    rq_activate_all_grippers(True)
    # end: URCap Program Node
  end
  $ 60 "zero_ftsensor()"
  zero_ftsensor()
  $ 61 "EXTT"
  $ 62 "Set GRP_3F_Enable=Off"
  set_standard_digital_out(4, False)
  $ 63 "Set BarcodeTrigger=Off"
  set_standard_digital_out(6, False)
  $ 64 "Set GRP_3F_Decap=Off"
  set_standard_digital_out(3, False)
  $ 65 "Set GRP_3F_Cap=Off"
  set_standard_digital_out(2, False)
  $ 66 "Set GRP_3F_Open=Off"
  set_standard_digital_out(5, False)
  $ 67 "PSE_T≔get_tool_free_pose(dir=[0,0,0.150], move_in_base_frame=True)"
  global PSE_T=get_tool_free_pose(dir=[0,0,0.150], move_in_base_frame=True)
  $ 68 "If is_reachable(Base_const, [PSE_T])"
  if (is_reachable(p[0.0,0.0,0.0,0.0,0.0,0.0], [PSE_T])):
    $ 69 "MoveL"
    $ 70 "PSE_T" "breakAfter"
    movel(PSE_T, a=1.2, v=0.15)
  end
  $ 71 "powder dispensing variable init"
  $ 72 "Start_thread≔ False "
  global Start_thread=  False
  $ 73 "vib_thread≔ False "
  global vib_thread=  False
  $ 74 "kp≔0.0015"
  global kp=0.0015
  $ 75 "ki≔0.0001"
  global ki=0.0001
  $ 76 "kd≔0.01"
  global kd=0.01
  $ 77 "dt≔0.03"
  global dt=0.03
  $ 78 "Integral_error≔0"
  global Integral_error=0
  $ 79 "current_error≔0"
  global current_error=0
  $ 80 "previous_error≔0"
  global previous_error=0
  $ 81 "tilt_increment≔0"
  global tilt_increment=0
  $ 82 "tilt_angle≔0"
  global tilt_angle=0
  $ 83 "diff≔0"
  global diff=0
  $ 84 "current_pose≔get_actual_tcp_pose()"
  global current_pose= get_actual_tcp_pose ()
  $ 85 "Relative_trans≔p[0, 0, -0.035, 0, 0, 0]"
  global Relative_trans=p[0, 0, -0.035, 0, 0, 0]
  $ 86 "ContA_plc_offst≔p[-0.00205, 0.02547, 0.03730, -0.03, -2.183, 6.165]"
  global ContA_plc_offst=p[-0.00205, 0.02547, 0.03730, -0.03, -2.183, 6.165]
  $ 87 "PowA_50_offset≔p[0.21808, -0.19943, 0.06584, 0, 0, 0]"
  global PowA_50_offset=p[0.21808, -0.19943, 0.06584, 0, 0, 0]
  $ 89 "tilt_init_reference()"
  tilt_init_reference()
  $ 90 "switch_spat_M≔ True "
  global switch_spat_M=  True
  $ 91 "switch_spat_S≔ True "
  global switch_spat_S=  True
  $ 92 "switch_spat_F_M≔ True "
  global switch_spat_F_M=  True
  $ 93 "switch_spat_F_S≔ True "
  global switch_spat_F_S=  True
  $ 94 "last_scale≔0"
  global last_scale=0
  $ 95 "W_EMPTY≔51.3"
  global W_EMPTY=51.3
  $ 768 "Thread_1"
  thread Thread_1():
    while (True):
      $ 769 "If Start_thread≟ True "
      if (Start_thread ==   True  ):
        $ 770 "weight_value≔get_weight()"
        global weight_value=get_weight()
        $ 771 "Wait: 0.1"
        sleep(0.1)
        $ 772 "sync()"
        sync()
      end
      $ 773 "sync()"
      sync()
    end
  end
  threadId_Thread_1 = run Thread_1()
  $ 774 "Thread_2"
  thread Thread_2():
    while (True):
      $ 775 "Loop vib_thread≟ True "
      thread Thread_while_775():
        while (True):
          $ 776 "diff≔target_weight-weight_value"
          global diff=target_weight-weight_value
          $ 777 "If diff>0.02 and spatula≠'spatula_flat_S'"
          global thread_flag_777=0
          thread Thread_if_777():
            $ 779 "Set AO[0]=4.0"
            set_standard_analog_out(0, 0.4)
            thread_flag_777 = 1
          end
          if (diff>0.02  and  spatula != "spatula_flat_S"):
            global thread_handler_777=run Thread_if_777()
            while (thread_flag_777 == 0):
              if not(diff>0.02  and  spatula != "spatula_flat_S"):
                kill thread_handler_777
                thread_flag_777 = 2
              else:
                sync()
              end
            end
          else:
            thread_flag_777 = 2
          end
          if (thread_flag_777 == 2):
            $ 780 "ElseIf diff>0.02 and spatula≟'spatula_flat_S'"
            if (diff>0.02 and spatula == "spatula_flat_S"):
              $ 781 "vibration_3()"
              vibration_3()
            else:
              $ 782 "ElseIf diff≤0.03"
              global thread_flag_782=0
              thread Thread_if_782():
                $ 783 "vibration_2()"
                vibration_2()
                thread_flag_782 = 1
              end
              if (diff <= 0.03):
                global thread_handler_782=run Thread_if_782()
                while (thread_flag_782 == 0):
                  if not(diff <= 0.03):
                    kill thread_handler_782
                    thread_flag_782 = 2
                  else:
                    sync()
                  end
                end
              else:
                thread_flag_782 = 2
              end
              if (thread_flag_782 == 2):
                $ 788 "Else" "noBreak"
                $ 789 "Set AO[0]=0.0"
                set_standard_analog_out(0, 0.0)
              end
            end
          end
        end
      end
      if (vib_thread ==   True  ):
        global thread_handler_775=run Thread_while_775()
        while (vib_thread ==   True  ):
          sync()
        end
        kill thread_handler_775
      end
      $ 790 "sync()"
      sync()
    end
  end
  threadId_Thread_2 = run Thread_2()
  while (True):
    $ 96 "Robot Program"
    $ 97 "MAIN"
    $ 98 "command_manager(external_control='uGO', cond_suspend=(ITM_Manipulated and AMR_AtTarget and AMR_Charging and AMR_Battery<40), cond_unsuspend=(AMR_Battery≟60))"
    command_manager(external_control="uGO", cond_suspend=(ITM_Manipulated  and  AMR_AtTarget  and  AMR_Charging  and  AMR_Battery<40), cond_unsuspend=(AMR_Battery == 60))
    $ 99 "log_state(STATE_Info)"
    log_state(STATE_Info)
    $ 100 "Switch STATE"
    switch_1 = STATE
    $ 101 "Case 1"
    if (1 == switch_1):
      $ 102 "Stopping"
      $ 103 "STATE_Info≔'Stopping'"
      global STATE_Info="Stopping"
      $ 104 "end_freedrive_mode()"
      end_freedrive_mode()
      $ 105 "Set"
      set_tcp(p[0.0,0.0,0.161,3.1415,0.0,0.0])
      $ 106 "PSE_T≔get_tool_free_pose(dir=[0,0,0.150], move_in_base_frame=True)"
      global PSE_T=get_tool_free_pose(dir=[0,0,0.150], move_in_base_frame=True)
      $ 107 "If is_reachable(Base_const, [PSE_T])"
      if (is_reachable(p[0.0,0.0,0.0,0.0,0.0,0.0], [PSE_T])):
        $ 108 "MoveL"
        $ 109 "PSE_T" "breakAfter"
        movel(PSE_T, a=1.2, v=0.15)
      end
      $ 110 "do_transition(keep_rxry=OBJ_Picked, r=0)"
      do_transition(keep_rxry=OBJ_Picked, r=0)
      $ 119 "Call Sub_AMR_MiR_V3"
      Sub_AMR_MiR_V3()
      $ 120 "If stopping() and AMR_Done"
      if (stopping()  and  AMR_Done):
        $ 121 "STATE≔2"
        global STATE=2
        $ 122 "ugo_update_outputs()"
        ugo_update_outputs()
      end
    elif (2 == switch_1):
      $ 123 "Case 2"
      $ 124 "Stopped"
      $ 125 "STATE_Info≔'Stopped'"
      global STATE_Info="Stopped"
      $ 126 "Call Sub_AMR_MiR_V3"
      Sub_AMR_MiR_V3()
      $ 127 "If CMD_Reset  or PB_Start"
      if (CMD_Reset   or  get_standard_digital_in(0)):
        $ 128 "STATE≔3"
        global STATE=3
        $ 129 "ugo_update_outputs()"
        ugo_update_outputs()
      end
    elif (3 == switch_1):
      $ 130 "Case 3"
      $ 131 " Resetting"
      $ 132 "STATE_Info≔'Resetting'"
      global STATE_Info="Resetting"
      $ 133 "uML"
      $ 134 "reset_error()"
      reset_error()
      $ 135 "reset_warning()"
      reset_warning()
      $ 136 "PROCESS_Step≔0"
      global PROCESS_Step=0
      $ 137 "PROCESS_Info≔''"
      global PROCESS_Info=""
      $ 138 "ARM_Referenced≔ False "
      global ARM_Referenced=  False
      $ 139 "WRK_Done≔ False "
      global WRK_Done=  False
      $ 140 "ITM_Prepared≔ False "
      global ITM_Prepared=  False
      $ 141 "ITM_Manipulated≔ False "
      global ITM_Manipulated=  False
      $ 142 "STP≔0"
      global STP=0
      $ 143 "Action≔0"
      global Action=0
      $ 144 "Action_Info≔''"
      global Action_Info=""
      $ 145 "ITM_ID≔0"
      global ITM_ID=0
      $ 146 "JIG≔0"
      global JIG=0
      $ 147 "JIG_Slot≔0"
      global JIG_Slot=0
      $ 148 "Task_info≔''"
      global Task_info=""
      $ 149 "Set"
      set_tcp(p[0.0,0.0,0.161,3.1415,0.0,0.0])
      $ 150 "App"
      $ 151 "'ADD APPLICATION SPECIFIC COMMANDS'"
      # 'ADD APPLICATION SPECIFIC COMMANDS'
      $ 152 "OBJ_Type≔0"
      global OBJ_Type=0
      $ 153 "OBJ_Nbr≔0"
      global OBJ_Nbr=0
      $ 154 "If CNT_Rack_Output≥50"
      if (CNT_Rack_Output >= 50):
        $ 155 "CNT_Rack_Output≔0"
        global CNT_Rack_Output=0
      end
      $ 156 "TASK≔struct(ID=0, NAVI=struct(target=0, footprint=0, protectiveOff=0, dock=0), WORK=struct(ITM_ID_Src=0, JIG_ID_Src=0, OBJ_Nbr_Src=0, ACT_Src=0, ITM_ID_Tgt=0, JIG_ID_Tgt=0, OBJ_Nbr_Tgt=0, ACT_Tgt=0, OBJ_Type=0))"
      global TASK=struct(ID=0, NAVI=struct(target=0, footprint=0, protectiveOff=0, dock=0), WORK=struct(ITM_ID_Src=0, JIG_ID_Src=0, OBJ_Nbr_Src=0, ACT_Src=0, ITM_ID_Tgt=0, JIG_ID_Tgt=0, OBJ_Nbr_Tgt=0, ACT_Tgt=0, OBJ_Type=0))
      $ 157 "Call Sub_AMR_MiR_V3"
      Sub_AMR_MiR_V3()
      $ 158 "If resetting() and AMR_Done"
      if (resetting()  and  AMR_Done):
        $ 159 "STATE≔4"
        global STATE=4
        $ 160 "ugo_update_outputs()"
        ugo_update_outputs()
      end
    elif (4 == switch_1):
      $ 161 "Case 4"
      $ 162 "Idle"
      $ 163 "STATE_Info≔'Idle'"
      global STATE_Info="Idle"
      $ 164 "If CMD_Start"
      if (CMD_Start):
        $ 165 "STATE≔5"
        global STATE=5
        $ 166 "ugo_update_outputs()"
        ugo_update_outputs()
      end
    elif (5 == switch_1):
      $ 167 "Case 5"
      $ 168 "Starting"
      $ 169 "STATE_Info≔'Starting'"
      global STATE_Info="Starting"
      $ 170 "'ADD COMMANDS WHAT TO START WITH'"
      # 'ADD COMMANDS WHAT TO START WITH'
      $ 171 "Call Sub_AMR_MiR_V3"
      Sub_AMR_MiR_V3()
      $ 172 "get ugo data"
      $ 173 "Assign Tasks"
      $ 174 "TASK.ID = ugo_get_task()"
      TASK.ID = ugo_get_task()
      $ 175 "If TASK.ID≟1"
      if (TASK.ID == 1):
        $ 176 "Task_info≔'Charge'"
        global Task_info="Charge"
        $ 177 "Parameters"
        $ 178 "AMR_PosTarget≔1"
        global AMR_PosTarget=1
      else:
        $ 179 "ElseIf TASK.ID≟9"
        if (TASK.ID == 9):
          $ 180 "'Pick Sarstedt Rack from Variable source'"
          # 'Pick Sarstedt Rack from Variable source'
          $ 181 "Task_info≔'Navigate to Target'"
          global Task_info="Navigate to Target"
          $ 182 "Parameters"
          $ 183 "AMR_PosTarget≔UGO.read_input('00','ITM_ID')"
          global AMR_PosTarget=UGO.read_input("00","ITM_ID")
        else:
          $ 184 "ElseIf TASK.ID≟49"
          if (TASK.ID == 49):
            $ 185 "Task_info≔'Pick Containers'"
            global Task_info="Pick Containers"
            $ 186 "Parameters"
            $ 187 "ITM_ID≔1"
            global ITM_ID=1
            $ 188 "OBJ_Type≔6"
            global OBJ_Type=6
            $ 189 "JIG≔15"
            global JIG=15
            $ 190 "AMR_PosTarget≔3"
            global AMR_PosTarget=3
          else:
            $ 191 "ElseIf TASK.ID≟50"
            if (TASK.ID == 50):
              $ 192 "Task_info≔'Decap Containers'"
              global Task_info="Decap Containers"
              $ 193 "Parameters"
              $ 194 "ITM_ID≔1"
              global ITM_ID=1
              $ 195 "OBJ_Type≔6"
              global OBJ_Type=6
              $ 196 "JIG≔16"
              global JIG=16
              $ 197 "AMR_PosTarget≔5"
              global AMR_PosTarget=5
            else:
              $ 198 "ElseIf TASK.ID≟51"
              if (TASK.ID == 51):
                $ 199 "Task_info≔'Detect Spatula and transfer powder'"
                global Task_info="Detect Spatula and transfer powder"
                $ 200 "Parameters"
                $ 201 "ITM_ID≔1"
                global ITM_ID=1
                $ 202 "target_weight≔(UGO.read_input('00','Target_weight'))/1000"
                global target_weight=(UGO.read_input("00","Target_weight"))/1000
                $ 203 "OBJ_Type≔8"
                global OBJ_Type=8
                $ 204 "JIG≔16"
                global JIG=16
                $ 205 "AMR_PosTarget≔5"
                global AMR_PosTarget=5
              else:
                $ 206 "ElseIf TASK.ID≟52"
                if (TASK.ID == 52):
                  $ 207 "Task_info≔'Pick Powder'"
                  global Task_info="Pick Powder"
                  $ 208 "Parameters"
                  $ 209 "ITM_ID≔1"
                  global ITM_ID=1
                  $ 210 "OBJ_Type≔6"
                  global OBJ_Type=6
                  $ 211 "JIG≔15"
                  global JIG=15
                  $ 212 "AMR_PosTarget≔3"
                  global AMR_PosTarget=3
                else:
                  $ 213 "ElseIf TASK.ID≟53"
                  if (TASK.ID == 53):
                    $ 214 "Task_info≔'Decap Powder'"
                    global Task_info="Decap Powder"
                    $ 215 "Parameters"
                    $ 216 "ITM_ID≔1"
                    global ITM_ID=1
                    $ 217 "OBJ_Type≔6"
                    global OBJ_Type=6
                    $ 218 "JIG≔1"
                    global JIG=1
                    $ 219 "AMR_PosTarget≔5"
                    global AMR_PosTarget=5
                  else:
                    $ 220 "ElseIf TASK.ID≟54"
                    if (TASK.ID == 54):
                      $ 221 "Task_info≔'Empty and swap Powder container'"
                      global Task_info="Empty and swap Powder container"
                      $ 230 "Parameters"
                      $ 231 "ITM_ID≔1"
                      global ITM_ID=1
                      $ 233 "W_now≔(UGO.read_input('00','Container_weight'))/1000"
                      global W_now=(UGO.read_input("00","Container_weight"))/1000
                      $ 234 "Pow_name≔(UGO.read_input('00','Powder_name'))"
                      global Pow_name=(UGO.read_input("00","Powder_name"))
                      $ 235 "scooping_init()"
                      scooping_init()
                      $ 236 "target_weight≔W_now-W_EMPTY-(0.002*W_FULL)"
                      global target_weight=W_now-W_EMPTY-(0.002*W_FULL)
                      $ 237 "OBJ_Type≔6"
                      global OBJ_Type=6
                      $ 238 "JIG≔17"
                      global JIG=17
                      $ 239 "AMR_PosTarget≔5"
                      global AMR_PosTarget=5
                    else:
                      $ 240 "ElseIf TASK.ID≟55"
                      if (TASK.ID == 55):
                        $ 241 "Task_info≔'Place Powder'"
                        global Task_info="Place Powder"
                        $ 242 "Parameters"
                        $ 243 "ITM_ID≔1"
                        global ITM_ID=1
                        $ 244 "OBJ_Type≔6"
                        global OBJ_Type=6
                        $ 245 "JIG≔21"
                        global JIG=21
                        $ 246 "AMR_PosTarget≔5"
                        global AMR_PosTarget=5
                      else:
                        $ 247 "ElseIf TASK.ID≟56"
                        if (TASK.ID == 56):
                          $ 248 "Task_info≔'Dose Powder'"
                          global Task_info="Dose Powder"
                          $ 249 "Parameters"
                          $ 250 "ITM_ID≔1"
                          global ITM_ID=1
                          $ 251 "target_weight≔(UGO.read_input('00','Target_weight'))/1000"
                          global target_weight=(UGO.read_input("00","Target_weight"))/1000
                          $ 252 "W_now≔(UGO.read_input('00','Container_weight'))/1000"
                          global W_now=(UGO.read_input("00","Container_weight"))/1000
                          $ 254 "Pow_name≔(UGO.read_input('00','Powder_name'))"
                          global Pow_name=(UGO.read_input("00","Powder_name"))
                          $ 255 "OBJ_Type≔6"
                          global OBJ_Type=6
                          $ 256 "JIG≔17"
                          global JIG=17
                          $ 257 "AMR_PosTarget≔5"
                          global AMR_PosTarget=5
                        else:
                          $ 258 "ElseIf TASK.ID≟57"
                          if (TASK.ID == 57):
                            $ 259 "Task_info≔'Recipe Powder dosing'"
                            global Task_info="Recipe Powder dosing"
                            $ 260 "Parameters"
                            $ 261 "ITM_ID≔1"
                            global ITM_ID=1
                            $ 262 "Pow_A≔(UGO.read_input('00','PowderA'))"
                            global Pow_A=(UGO.read_input("00","PowderA"))
                            $ 263 "Pow_B≔(UGO.read_input('00','PowderB'))"
                            global Pow_B=(UGO.read_input("00","PowderB"))
                            $ 264 "Pow_C≔(UGO.read_input('00','PowderC'))"
                            global Pow_C=(UGO.read_input("00","PowderC"))
                            $ 265 "Total_weight≔(UGO.read_input('00','Total_weight'))/1000"
                            global Total_weight=(UGO.read_input("00","Total_weight"))/1000
                            $ 266 "Pow_A_percent≔(UGO.read_input('00','PowderA_percentage'))/100"
                            global Pow_A_percent=(UGO.read_input("00","PowderA_percentage"))/100
                            $ 267 "Pow_B_percent≔(UGO.read_input('00','PowderB_percentage'))/100"
                            global Pow_B_percent=(UGO.read_input("00","PowderB_percentage"))/100
                            $ 268 "Pow_C_percent≔(UGO.read_input('00','PowderC_percentage'))/100"
                            global Pow_C_percent=(UGO.read_input("00","PowderC_percentage"))/100
                            $ 269 "OBJ_Type≔6"
                            global OBJ_Type=6
                            $ 270 "JIG≔17"
                            global JIG=17
                            $ 271 "AMR_PosTarget≔5"
                            global AMR_PosTarget=5
                          else:
                            $ 272 "ElseIf TASK.ID≟58"
                            if (TASK.ID == 58):
                              $ 273 "Task_info≔'Pick Powder containers'"
                              global Task_info="Pick Powder containers"
                              $ 274 "Parameters"
                              $ 275 "ITM_ID≔1"
                              global ITM_ID=1
                              $ 276 "OBJ_Type≔6"
                              global OBJ_Type=6
                              $ 277 "JIG≔15"
                              global JIG=15
                              $ 278 "AMR_PosTarget≔3"
                              global AMR_PosTarget=3
                            else:
                              $ 279 "Else" "noBreak"
                              $ 280 "set_error(ERROR_WRONG_ORDER)"
                              set_error(ERROR_WRONG_ORDER)
                            end
                          end
                        end
                      end
                    end
                  end
                end
              end
            end
          end
        end
      end
      $ 281 "test ugo"
      $ 282 "Wait: 0.2"
      sleep(0.2)
      $ 283 "ugo_update_outputs()"
      ugo_update_outputs()
      $ 284 "If starting() and AMR_Done"
      if (starting()  and  AMR_Done):
        $ 285 "log_message(Task_info, 'New Task: ')"
        log_message(Task_info, "New Task: ")
        $ 286 "log_message(to_str(TASK.ID), 'Task_ID: ')"
        log_message(to_str(TASK.ID), "Task_ID: ")
        $ 287 "do_transition(keep_rxry=OBJ_Picked)"
        do_transition(keep_rxry=OBJ_Picked)
        $ 288 "STATE≔6"
        global STATE=6
        $ 289 "ugo_update_outputs()"
        ugo_update_outputs()
      end
    elif (6 == switch_1):
      $ 290 "Case 6"
      $ 291 "Execute"
      $ 292 "STATE_Info≔'Execute'"
      global STATE_Info="Execute"
      $ 293 "If  not CMD_Hold and not CMD_Suspend"
      global thread_flag_293=0
      thread Thread_if_293():
        $ 294 "Switch PROCESS_Step"
        switch_2 = PROCESS_Step
        $ 295 "Case 0"
        if (0 == switch_2):
          $ 296 "PROCESS_Info≔'process control'"
          global PROCESS_Info="process control"
          $ 297 "log_process(PROCESS_Info)"
          log_process(PROCESS_Info)
          $ 298 "process control"
          $ 299 "If  not AMR_AtTarget"
          if (  not  AMR_AtTarget):
            $ 300 "PROCESS_Step≔1"
            global PROCESS_Step=1
          else:
            $ 301 "ElseIf (( not ITM_Prepared and  not WRK_Done) or (ITM_Prepared and WRK_Done))"
            if (((  not  ITM_Prepared  and    not  WRK_Done)  or  (ITM_Prepared  and  WRK_Done))):
              $ 302 "PROCESS_Step≔2"
              global PROCESS_Step=2
            else:
              $ 303 "ElseIf  not WRK_Done"
              if (  not  WRK_Done):
                $ 304 "PROCESS_Step≔3"
                global PROCESS_Step=3
              else:
                $ 305 "Else" "noBreak"
                $ 306 "task finished"
                $ 307 "PROCESS_Info≔''"
                global PROCESS_Info=""
                $ 308 "STATE≔7"
                global STATE=7
                $ 309 "ugo_update_outputs()"
                ugo_update_outputs()
              end
            end
          end
        elif (1 == switch_2):
          $ 310 "Case 1"
          $ 311 "navigate"
          $ 312 "'MOVING THE uML'"
          # 'MOVING THE uML'
          $ 313 "PROCESS_Info≔'move to target'"
          global PROCESS_Info="move to target"
          $ 314 "log_process(PROCESS_Info)"
          log_process(PROCESS_Info)
          $ 315 "If TASK.ID≟1"
          if (TASK.ID == 1):
            $ 316 "Action≔51"
            global Action=51
          else:
            $ 317 "Else" "noBreak"
            $ 318 "Action≔52"
            global Action=52
          end
          $ 319 "Call Sub_AMR_MiR_V3"
          Sub_AMR_MiR_V3()
          $ 320 "If AMR_Done"
          if (AMR_Done):
            $ 321 "PROCESS_Step≔0"
            global PROCESS_Step=0
          end
        elif (2 == switch_2):
          $ 322 "Case 2"
          $ 323 "prepare"
          $ 324 "'THINGS THAT HAVE TO BE DONE ONCE IN A SEQUENCE,WORKFLOW'"
          # 'THINGS THAT HAVE TO BE DONE ONCE IN A SEQUENCE,WORKFLOW'
          $ 325 "PROCESS_Info≔'prepare for work'"
          global PROCESS_Info="prepare for work"
          $ 326 "log_process(PROCESS_Info)"
          log_process(PROCESS_Info)
          $ 327 "If TASK.WORK.ITM_ID_Src>1"
          if (TASK.WORK.ITM_ID_Src>1):
            $ 328 "ITM_ID≔TASK.WORK.ITM_ID_Src"
            global ITM_ID=TASK.WORK.ITM_ID_Src
          else:
            $ 329 "ElseIf TASK.WORK.ITM_ID_Tgt>1"
            if (TASK.WORK.ITM_ID_Tgt>1):
              $ 330 "ITM_ID≔TASK.WORK.ITM_ID_Tgt"
              global ITM_ID=TASK.WORK.ITM_ID_Tgt
            end
          end
          $ 331 "If  not ARM_Referenced and (ITM_ID≠0)"
          if (  not  ARM_Referenced  and  (ITM_ID != 0)):
            $ 332 "STP≔1"
            global STP=1
          else:
            $ 333 "ElseIf ARM_Referenced or (ITM_ID≟0)"
            if (ARM_Referenced  or  (ITM_ID == 0)):
              $ 334 "STP≔2"
              global STP=2
            end
          end
          $ 335 "Switch STP"
          switch_3 = STP
          $ 336 "Case 1"
          if (1 == switch_3):
            $ 337 "reference"
            $ 338 "STP_Info≔'reference at target position'"
            global STP_Info="reference at target position"
            $ 339 "log_step(STP_Info)"
            log_step(STP_Info)
            $ 340 "If ITM_ID≟1"
            if (ITM_ID == 1):
              $ 341 "CAM_Done≔ True "
              global CAM_Done=  True
            else:
              $ 342 "Else" "noBreak"
              $ 343 "Action≔131"
              global Action=131
              $ 344 "Call Sub_Vision_V18"
              Sub_Vision_V18()
            end
            $ 346 "If CAM_Done and  not ERROR.FLAG"
            if (CAM_Done  and    not  ERROR.FLAG):
              $ 347 "log_step('ARM referenced')"
              log_step("ARM referenced")
              $ 348 "ARM_Referenced≔ True "
              global ARM_Referenced=  True
            end
          elif (2 == switch_3):
            $ 349 "Case 2"
            $ 350 "manipulate"
            $ 351 "STP_Info≔'manipulate item'"
            global STP_Info="manipulate item"
            $ 352 "log_step(STP_Info)"
            log_step(STP_Info)
            $ 353 "'In case pressing button is needed'"
            # 'In case pressing button is needed'
            $ 354 "If found_in_list(ITM_ID, ITM_ID_List)"
            if (found_in_list(ITM_ID, ITM_ID_List)):
              $ 355 "Switch ITM_ID"
              switch_4 = ITM_ID
              $ 356 "Case 0"
              if (0 == switch_4):
                $ 357 "ITM_Manipulated≔ not ITM_Manipulated"
                global ITM_Manipulated=  not  ITM_Manipulated
              elif (1 == switch_4):
                $ 358 "Case 1"
                $ 359 "ITM_Manipulated≔ not ITM_Manipulated"
                global ITM_Manipulated=  not  ITM_Manipulated
              elif (2 == switch_4):
                $ 360 "Case 2"
              else:
                $ 370 "Default Case"
                $ 371 "ITM_Manipulated≔ not ITM_Manipulated"
                global ITM_Manipulated=  not  ITM_Manipulated
              end
            end
          end
          $ 372 "ITM_Prepared≔(ITM_Manipulated or  not found_in_list(ITM_ID, ITM_ID_List)) and (ARM_Referenced or ITM_ID≟0) and  not WRK_Done"
          global ITM_Prepared=(ITM_Manipulated  or    not  found_in_list(ITM_ID, ITM_ID_List))  and  (ARM_Referenced  or  ITM_ID == 0)  and    not  WRK_Done
          $ 373 "STP≔0"
          global STP=0
          $ 374 "STP_Info≔''"
          global STP_Info=""
          $ 375 "PROCESS_Step≔0"
          global PROCESS_Step=0
        elif (3 == switch_2):
          $ 376 "Case 3"
          $ 377 "work"
          $ 378 "'ADD EVERY MACHINE, OBJECT, STATION TO WORK ON'"
          # 'ADD EVERY MACHINE, OBJECT, STATION TO WORK ON'
          $ 379 "Switch ITM_ID"
          switch_3 = ITM_ID
          $ 380 "Case 1"
          if (1 == switch_3):
            $ 381 "uLM"
            $ 382 "If TASK.ID≟12"
            if (TASK.ID == 12):
              $ 383 "fill racks"
              $ 384 "Action≔151"
              global Action=151
              $ 385 "Call Sub_Vision_V18"
              Sub_Vision_V18()
              $ 386 "If  not ERROR.FLAG"
              if (  not  ERROR.FLAG):
                $ 387 "Actions for the task"
                $ 388 "Action≔1"
                global Action=1
                $ 389 "JIG≔2"
                global JIG=2
                $ 390 "JIG_Slot≔CAM_Result[0]"
                global JIG_Slot=CAM_Result[0]
                $ 391 "OBJ_Nbr≔CAM_Result[0]"
                global OBJ_Nbr=CAM_Result[0]
                $ 392 "OBJ_Type≔2"
                global OBJ_Type=2
                $ 393 "Call Sub_Action_V4"
                Sub_Action_V4()
                $ 394 "If OBJ_Picked"
                if (OBJ_Picked):
                  $ 395 "CAM_Result.remove(0)"
                  CAM_Result.remove(0)
                  $ 396 "PRC_TubCounter≔PRC_TubCounter+1"
                  global PRC_TubCounter=PRC_TubCounter+1
                  $ 397 "If PRC_TubCounter%4≟0"
                  if (PRC_TubCounter%4 == 0):
                    $ 398 "JIG_Slot≔4"
                    global JIG_Slot=4
                  else:
                    $ 399 "Else" "noBreak"
                    $ 400 "JIG_Slot≔PRC_TubCounter%4"
                    global JIG_Slot=PRC_TubCounter%4
                  end
                  $ 401 "OBJ_Nbr≔ceil(PRC_TubCounter/4)"
                  global OBJ_Nbr=ceil(PRC_TubCounter/4)
                  $ 402 "Action≔2"
                  global Action=2
                  $ 403 "JIG≔4"
                  global JIG=4
                  $ 404 "Call Sub_Action_V4"
                  Sub_Action_V4()
                  $ 405 "Action≔151"
                  global Action=151
                  $ 406 "Call Sub_Vision_V18"
                  Sub_Vision_V18()
                end
              end
              $ 407 "If (CAM_Captures≥CAM_PRM_Retries) or (PRC_TubCounter≥32)"
              if ((CAM_Captures >= CAM_PRM_Retries)  or  (PRC_TubCounter >= 32)):
                $ 408 "PROCESS_Step≔0"
                global PROCESS_Step=0
                $ 409 "WRK_Done≔ True "
                global WRK_Done=  True
              end
            else:
              $ 410 "ElseIf TASK.ID≟49"
              if (TASK.ID == 49):
                $ 411 "Pick Powder container"
                $ 412 "Action≔131"
                global Action=131
                $ 413 "Call Sub_Vision_V18"
                Sub_Vision_V18()
                $ 414 "Action≔35"
                global Action=35
                $ 415 "Call Sub_Action_V4"
                Sub_Action_V4()
                $ 416 "PROCESS_Step≔0"
                global PROCESS_Step=0
                $ 417 "WRK_Done≔ True "
                global WRK_Done=  True
              else:
                $ 418 "ElseIf TASK.ID≟50"
                if (TASK.ID == 50):
                  $ 419 "Decap containers"
                  $ 420 "Action≔36"
                  global Action=36
                  $ 421 "Call Sub_Action_V4"
                  Sub_Action_V4()
                  $ 422 "PROCESS_Step≔0"
                  global PROCESS_Step=0
                  $ 423 "WRK_Done≔ True "
                  global WRK_Done=  True
                else:
                  $ 424 "ElseIf TASK.ID≟51"
                  if (TASK.ID == 51):
                    $ 425 "Detect Spatula and transfer powder"
                    $ 426 "Action≔131"
                    global Action=131
                    $ 427 "Call Sub_Vision_V18"
                    Sub_Vision_V18()
                    $ 428 "Action≔37"
                    global Action=37
                    $ 429 "Call Sub_Action_V4"
                    Sub_Action_V4()
                    $ 430 "PROCESS_Step≔0"
                    global PROCESS_Step=0
                    $ 431 "WRK_Done≔ True "
                    global WRK_Done=  True
                  else:
                    $ 432 "ElseIf TASK.ID≟52"
                    if (TASK.ID == 52):
                      $ 433 "Pick Powder container"
                      $ 434 "Action≔131"
                      global Action=131
                      $ 435 "Call Sub_Vision_V18"
                      Sub_Vision_V18()
                      $ 436 "Action≔39"
                      global Action=39
                      $ 437 "Call Sub_Action_V4"
                      Sub_Action_V4()
                      $ 438 "PROCESS_Step≔0"
                      global PROCESS_Step=0
                      $ 439 "WRK_Done≔ True "
                      global WRK_Done=  True
                    else:
                      $ 440 "ElseIf TASK.ID≟53"
                      if (TASK.ID == 53):
                        $ 441 "Decap containerA"
                        $ 442 "Action≔40"
                        global Action=40
                        $ 443 "Call Sub_Action_V4"
                        Sub_Action_V4()
                        $ 444 "PROCESS_Step≔0"
                        global PROCESS_Step=0
                        $ 445 "WRK_Done≔ True "
                        global WRK_Done=  True
                      else:
                        $ 446 "ElseIf TASK.ID≟55"
                        if (TASK.ID == 55):
                          $ 447 "Place Powder"
                          $ 448 "Action≔131"
                          global Action=131
                          $ 449 "Call Sub_Vision_V18"
                          Sub_Vision_V18()
                          $ 450 "Action≔41"
                          global Action=41
                          $ 451 "Call Sub_Action_V4"
                          Sub_Action_V4()
                          $ 452 "PROCESS_Step≔0"
                          global PROCESS_Step=0
                          $ 453 "WRK_Done≔ True "
                          global WRK_Done=  True
                        else:
                          $ 454 "ElseIf TASK.ID≟54"
                          if (TASK.ID == 54):
                            $ 455 "Empty and swap container"
                            $ 456 "Action≔131"
                            global Action=131
                            $ 457 "Call Sub_Vision_V18"
                            Sub_Vision_V18()
                            $ 458 "Action≔42"
                            global Action=42
                            $ 459 "Call Sub_Action_V4"
                            Sub_Action_V4()
                            $ 460 "PROCESS_Step≔0"
                            global PROCESS_Step=0
                            $ 461 "WRK_Done≔ True "
                            global WRK_Done=  True
                          else:
                            $ 462 "ElseIf TASK.ID≟56"
                            if (TASK.ID == 56):
                              $ 463 "Dispense Powder"
                              $ 464 "Action≔131"
                              global Action=131
                              $ 465 "Call Sub_Vision_V18"
                              Sub_Vision_V18()
                              $ 466 "Action≔43"
                              global Action=43
                              $ 467 "Call Sub_Action_V4"
                              Sub_Action_V4()
                              $ 468 "PROCESS_Step≔0"
                              global PROCESS_Step=0
                              $ 469 "WRK_Done≔ True "
                              global WRK_Done=  True
                            else:
                              $ 470 "ElseIf TASK.ID≟57"
                              if (TASK.ID == 57):
                                $ 471 "Recipe Dosing"
                                $ 472 "Action≔48"
                                global Action=48
                                $ 473 "Call Sub_Action_V4"
                                Sub_Action_V4()
                                $ 474 "recipe_init(Pow_A, Pow_B, Pow_C, Total_weight, Pow_A_percent, Pow_B_percent, Pow_C_percent)"
                                recipe_init(Pow_A, Pow_B, Pow_C, Total_weight, Pow_A_percent, Pow_B_percent, Pow_C_percent)
                                $ 475 "Loop recipe_next()≟ True "
                                while (recipe_next() ==   True  ):
                                  $ 476 "Action≔44"
                                  global Action=44
                                  $ 477 "Call Sub_Action_V4"
                                  Sub_Action_V4()
                                  $ 478 "JIG≔21"
                                  global JIG=21
                                  $ 479 "Action≔131"
                                  global Action=131
                                  $ 480 "Call Sub_Vision_V18"
                                  Sub_Vision_V18()
                                  $ 481 "Action≔45"
                                  global Action=45
                                  $ 482 "Call Sub_Action_V4"
                                  Sub_Action_V4()
                                  $ 483 "dosing_start()"
                                  dosing_start()
                                  $ 484 "JIG≔17"
                                  global JIG=17
                                  $ 485 "Action≔131"
                                  global Action=131
                                  $ 486 "Call Sub_Vision_V18"
                                  Sub_Vision_V18()
                                  $ 487 "Action≔46"
                                  global Action=46
                                  $ 488 "Call Sub_Action_V4"
                                  Sub_Action_V4()
                                  $ 489 "dosing_end()"
                                  dosing_end()
                                end
                                $ 490 "PROCESS_Step≔0"
                                global PROCESS_Step=0
                                $ 491 "WRK_Done≔ True "
                                global WRK_Done=  True
                              else:
                                $ 492 "ElseIf TASK.ID≟58"
                                if (TASK.ID == 58):
                                  $ 493 "Pick Powder containers"
                                  $ 494 "Num_cont_picked≔0"
                                  global Num_cont_picked=0
                                  $ 495 "powder_position≔'Position1'"
                                  global powder_position="Position1"
                                  $ 496 "Loop Num_cont_picked<3"
                                  while (Num_cont_picked<3):
                                    $ 497 "Action≔131"
                                    global Action=131
                                    $ 498 "Call Sub_Vision_V18"
                                    Sub_Vision_V18()
                                    $ 499 "Action≔47"
                                    global Action=47
                                    $ 500 "Call Sub_Action_V4"
                                    Sub_Action_V4()
                                  end
                                  $ 501 "PROCESS_Step≔0"
                                  global PROCESS_Step=0
                                  $ 502 "WRK_Done≔ True "
                                  global WRK_Done=  True
                                end
                              end
                            end
                          end
                        end
                      end
                    end
                  end
                end
              end
            end
          elif (2 == switch_3):
            $ 503 "Case 2"
          elif (5 == switch_3):
            $ 545 "Case 5"
          elif (20 == switch_3):
            $ 553 "Case 20"
          elif (43 == switch_3):
            $ 615 "Case 43"
          else:
            $ 623 "Default Case"
            $ 624 "WRK_Done≔ True "
            global WRK_Done=  True
            $ 625 "PROCESS_Step≔0"
            global PROCESS_Step=0
          end
        end
        thread_flag_293 = 1
      end
      if (  not  CMD_Hold and not CMD_Suspend):
        global thread_handler_293=run Thread_if_293()
        while (thread_flag_293 == 0):
          if not(  not  CMD_Hold and not CMD_Suspend):
            kill thread_handler_293
            thread_flag_293 = 2
          else:
            sync()
          end
        end
      else:
        thread_flag_293 = 2
      end
      $ 626 "If CMD_Hold"
      if (CMD_Hold):
        $ 627 "STATE≔9"
        global STATE=9
        $ 628 "ugo_update_outputs()"
        ugo_update_outputs()
      else:
        $ 629 "ElseIf CMD_Suspend"
        if (CMD_Suspend):
          $ 630 "STATE≔12"
          global STATE=12
          $ 631 "ugo_update_outputs()"
          ugo_update_outputs()
        end
      end
    elif (7 == switch_1):
      $ 632 "Case 7"
      $ 633 "Completing"
      $ 634 "STATE_Info≔'Completing'"
      global STATE_Info="Completing"
      $ 635 "'ADD COMMANDS FOR COMPLETING THE PROCESS'"
      # 'ADD COMMANDS FOR COMPLETING THE PROCESS'
      $ 636 "do_transition(keep_rxry=OBJ_Picked)"
      do_transition(keep_rxry=OBJ_Picked)
      $ 637 "Call Sub_AMR_MiR_V3"
      Sub_AMR_MiR_V3()
      $ 638 "If completing() and AMR_Done"
      if (completing()  and  AMR_Done):
        $ 639 "STATE≔8"
        global STATE=8
        $ 640 "ugo_update_outputs()"
        ugo_update_outputs()
      end
    elif (8 == switch_1):
      $ 641 "Case 8"
      $ 642 "Complete"
      $ 643 "STATE_Info≔'Complete'"
      global STATE_Info="Complete"
      $ 644 "If CMD_Reset"
      if (CMD_Reset):
        $ 645 "STATE≔3"
        global STATE=3
        $ 646 "ugo_update_outputs()"
        ugo_update_outputs()
      end
    elif (9 == switch_1):
      $ 647 "Case 9"
      $ 648 "Holding"
      $ 649 "STATE_Info≔'Holding'"
      global STATE_Info="Holding"
      $ 650 "stopl(0.5)"
      stopl(0.5)
      $ 651 "Call Sub_AMR_MiR_V3"
      Sub_AMR_MiR_V3()
      $ 652 "If holding() and AMR_Done"
      if (holding()  and  AMR_Done):
        $ 653 "STATE≔10"
        global STATE=10
        $ 654 "ugo_update_outputs()"
        ugo_update_outputs()
      end
    elif (10 == switch_1):
      $ 655 "Case 10"
      $ 656 "Held"
      $ 657 "STATE_Info≔'Held'"
      global STATE_Info="Held"
      $ 658 "If CMD_Unhold"
      if (CMD_Unhold):
        $ 659 "end_freedrive_mode()"
        end_freedrive_mode()
        $ 660 "STATE≔11"
        global STATE=11
        $ 661 "ugo_update_outputs()"
        ugo_update_outputs()
      else:
        $ 662 "ElseIf FNC_Freedrive"
        if (FNC_Freedrive):
          $ 663 "freedrive_mode()"
          freedrive_mode()
        else:
          $ 664 "Else" "noBreak"
          $ 665 "end_freedrive_mode()"
          end_freedrive_mode()
        end
      end
    elif (11 == switch_1):
      $ 666 "Case 11"
      $ 667 "Unholding"
      $ 668 "STATE_Info≔'Unholding'"
      global STATE_Info="Unholding"
      $ 669 "Clearing"
      $ 670 "Switch ERROR.ID"
      switch_2 = ERROR.ID
      $ 671 "Case 1002"
      if (1002 == switch_2):
        $ 672 "AMR_AtTarget≔ False "
        global AMR_AtTarget=  False
        $ 673 "ARM_Referenced≔ False "
        global ARM_Referenced=  False
        $ 674 "ITM_Prepared≔ False "
        global ITM_Prepared=  False
        $ 675 "PROCESS_Step≔1"
        global PROCESS_Step=1
      elif (2007 == switch_2):
        $ 676 "Case 2007"
        $ 677 "PROCESS_Step≔1"
        global PROCESS_Step=1
      end
      $ 678 "reset_error()"
      reset_error()
      $ 679 "reset_warning()"
      reset_warning()
      $ 680 "OBJ_Picked≔gripper_has_object()"
      global OBJ_Picked=gripper_has_object()
      $ 681 "Call Sub_AMR_MiR_V3"
      Sub_AMR_MiR_V3()
      $ 682 "If unholding() and AMR_Done"
      if (unholding()  and  AMR_Done):
        $ 683 "STATE≔6"
        global STATE=6
        $ 684 "ugo_update_outputs()"
        ugo_update_outputs()
      end
    elif (12 == switch_1):
      $ 685 "Case 12"
      $ 686 "Suspending"
      $ 687 "STATE_Info≔'Suspending'"
      global STATE_Info="Suspending"
      $ 688 "PROCESS_Info≔str_cat(PROCESS_Info, ' suspended')"
      global PROCESS_Info=str_cat(PROCESS_Info, " suspended")
      $ 689 "If suspending()"
      if (suspending()):
        $ 690 "STATE≔13"
        global STATE=13
        $ 691 "ugo_update_outputs()"
        ugo_update_outputs()
      end
    elif (13 == switch_1):
      $ 692 "Case 13"
      $ 693 "Suspended"
      $ 694 "STATE_Info≔'Suspended'"
      global STATE_Info="Suspended"
      $ 695 "Call Sub_AMR_MiR_V3"
      Sub_AMR_MiR_V3()
      $ 696 "If CMD_Unsuspend"
      if (CMD_Unsuspend):
        $ 697 "STATE≔14"
        global STATE=14
        $ 698 "ugo_update_outputs()"
        ugo_update_outputs()
      end
    elif (14 == switch_1):
      $ 699 "Case 14"
      $ 700 "Unsuspending"
      $ 701 "STATE_Info≔'Unsuspending'"
      global STATE_Info="Unsuspending"
      $ 702 "PROCESS_Step≔0"
      global PROCESS_Step=0
      $ 703 "If unsuspending()"
      if (unsuspending()):
        $ 704 "STATE≔6"
        global STATE=6
        $ 705 "ugo_update_outputs()"
        ugo_update_outputs()
      end
    elif (15 == switch_1):
      $ 706 "Case 15"
      $ 707 "Aborting"
      $ 708 "STATE_Info≔'Aborting'"
      global STATE_Info="Aborting"
      $ 709 "If aborting()"
      if (aborting()):
        $ 710 "STATE≔16"
        global STATE=16
        $ 711 "ugo_update_outputs()"
        ugo_update_outputs()
      end
    elif (16 == switch_1):
      $ 712 "Case 16"
      $ 713 "Aborted"
      $ 714 "STATE_Info≔'Aborted'"
      global STATE_Info="Aborted"
      $ 715 "If CMD_Clear"
      if (CMD_Clear):
        $ 716 "STATE≔17"
        global STATE=17
        $ 717 "ugo_update_outputs()"
        ugo_update_outputs()
      end
    elif (17 == switch_1):
      $ 718 "Case 17"
      $ 719 "Clearing"
      $ 720 "STATE_Info≔'Clearing'"
      global STATE_Info="Clearing"
      $ 721 "Clearing"
      $ 722 "reset_warning()"
      reset_warning()
      $ 723 "reset_error()"
      reset_error()
      $ 724 "If clearing()"
      if (clearing()):
        $ 725 "STATE≔2"
        global STATE=2
        $ 726 "ugo_update_outputs()"
        ugo_update_outputs()
      end
    end
    $ 727 "log_state(STATE_Info)"
    log_state(STATE_Info)
    $ 728 "log_warning(WARNING.MSG)"
    log_warning(WARNING.MSG)
    $ 729 "log_error(ERROR.MSG)"
    log_error(ERROR.MSG)
    $ 730 "Times"
    $ 731 "Switch STATE"
    switch_1 = STATE
    $ 732 "Case 1"
    if (1 == switch_1):
      $ 733 "TM_St_Stopping≔get_time(STATE_Times[STATE-1])"
      global TM_St_Stopping=get_time(STATE_Times[STATE-1])
    elif (2 == switch_1):
      $ 734 "Case 2"
      $ 735 "TM_St_Stopped≔get_time(STATE_Times[STATE-1])"
      global TM_St_Stopped=get_time(STATE_Times[STATE-1])
    elif (3 == switch_1):
      $ 736 "Case 3"
      $ 737 "TM_St_Resetting≔get_time(STATE_Times[STATE-1])"
      global TM_St_Resetting=get_time(STATE_Times[STATE-1])
    elif (4 == switch_1):
      $ 738 "Case 4"
      $ 739 "TM_St_Idle≔get_time(STATE_Times[STATE-1])"
      global TM_St_Idle=get_time(STATE_Times[STATE-1])
    elif (5 == switch_1):
      $ 740 "Case 5"
      $ 741 "TM_St_Starting≔get_time(STATE_Times[STATE-1])"
      global TM_St_Starting=get_time(STATE_Times[STATE-1])
    elif (6 == switch_1):
      $ 742 "Case 6"
      $ 743 "TM_St_Execute≔get_time(STATE_Times[STATE-1])"
      global TM_St_Execute=get_time(STATE_Times[STATE-1])
    elif (7 == switch_1):
      $ 744 "Case 7"
      $ 745 "TM_St_Completin≔get_time(STATE_Times[STATE-1])"
      global TM_St_Completin=get_time(STATE_Times[STATE-1])
    elif (8 == switch_1):
      $ 746 "Case 8"
      $ 747 "TM_St_Complete≔get_time(STATE_Times[STATE-1])"
      global TM_St_Complete=get_time(STATE_Times[STATE-1])
    elif (9 == switch_1):
      $ 748 "Case 9"
      $ 749 "TM_St_Holding≔get_time(STATE_Times[STATE-1])"
      global TM_St_Holding=get_time(STATE_Times[STATE-1])
    elif (10 == switch_1):
      $ 750 "Case 10"
      $ 751 "TM_St_Held≔get_time(STATE_Times[STATE-1])"
      global TM_St_Held=get_time(STATE_Times[STATE-1])
    elif (11 == switch_1):
      $ 752 "Case 11"
      $ 753 "TM_St_Unholding≔get_time(STATE_Times[STATE-1])"
      global TM_St_Unholding=get_time(STATE_Times[STATE-1])
    elif (12 == switch_1):
      $ 754 "Case 12"
      $ 755 "TM_St_Suspendin≔get_time(STATE_Times[STATE-1])"
      global TM_St_Suspendin=get_time(STATE_Times[STATE-1])
    elif (13 == switch_1):
      $ 756 "Case 13"
      $ 757 "TM_St_Suspended≔get_time(STATE_Times[STATE-1])"
      global TM_St_Suspended=get_time(STATE_Times[STATE-1])
    elif (14 == switch_1):
      $ 758 "Case 14"
      $ 759 "TM_St_Unsuspend≔get_time(STATE_Times[STATE-1])"
      global TM_St_Unsuspend=get_time(STATE_Times[STATE-1])
    elif (15 == switch_1):
      $ 760 "Case 15"
      $ 761 "TM_St_Aborting≔get_time(STATE_Times[STATE-1])"
      global TM_St_Aborting=get_time(STATE_Times[STATE-1])
    elif (16 == switch_1):
      $ 762 "Case 16"
      $ 763 "TM_St_Aborted≔get_time(STATE_Times[STATE-1])"
      global TM_St_Aborted=get_time(STATE_Times[STATE-1])
    elif (17 == switch_1):
      $ 764 "Case 17"
      $ 765 "TM_St_Clearing≔get_time(STATE_Times[STATE-1])"
      global TM_St_Clearing=get_time(STATE_Times[STATE-1])
    end
    $ 767 "Wait: 0.1"
    sleep(0.1)
  end
end
